Fanuc KAREL source: KA00148.KL

PROGRAM KA00148
%NOLOCKGROUP
VAR
  SRC: ARRAY[4] OF INTEGER
  DST: ARRAY[4] OF STRING[20]
BEGIN
  DST = SRC
END KA00148
